(*
SPDX-FileCopyrightText: © 2026 Oleksandr Tiutyk <trofimich@gmail.com>
SPDX-License-Identifier: MIT
License: https://opensource.org/license/mit
*)

(*!
<summary>Provides shared comparer instances and selects them by generic value category.</summary>
<description>
Returned comparer interfaces borrow instances stored in this program; callers do not own or release them.
Selection does not inspect, validate or convert operand data. Callers must supply live descriptors whose
representations satisfy the selected concrete comparer. OBJECT selects natural ordering through IComparable;
it does not select byte or address ordering. Dictionary/set equality lookup is independent of this catalogue.
</description>
*)

PROGRAM StandardComparers
VAR_OUTPUT
	BoolComparer : BoolComparer;
	SIntComparer : SIntComparer;
	USIntComparer : USIntComparer;
	IntComparer : IntComparer;
	UIntComparer : UIntComparer;
	DIntComparer : DIntComparer;
	UDIntComparer : UDIntComparer;
	LIntComparer : LIntComparer;
	ULIntComparer : ULIntComparer;
	RealComparer : RealComparer;
	LRealComparer : LRealComparer;		
	StringComparer : StringComparer;
	WStringComparer : WStringComparer;
	TimeComparer : TimeComparer;
	LTimeComparer : LTimeComparer;
	DateComparer : DateComparer;
	LDateComparer : LDateComparer;
	DateAndTimeComparer : DateAndTimeComparer;
	LDateAndTimeComparer : LDateAndTimeComparer;
	TimeOfDayComparer : TimeOfDayComparer;	
	LTimeOfDayComparer : LTimeOfDayComparer;	
	ByteArrayComparer : ByteArrayComparer;
	ObjectComparer : ObjectComparer;
	//! <summary>Shared comparer that orders descriptor storage addresses without reading stored pointer values.</summary>
	StorageAddressComparer : StorageAddressComparer;	
END_VAR
VAR
	{attribute 'hide'} 
	_ClassName : STRING := __POUNAME();
END_VAR

{attribute 'monitoring' := 'call'}
PROPERTY ClassName : REFERENCE TO STRING
GET
ClassName REF= _ClassName;
END_GET
END_PROPERTY

(*!
<summary>Returns the shared comparer selected for a generic value category.</summary>
<description>
The result borrows a catalogue instance and does not transfer ownership. No operands are inspected or
converted; compatibility and operand lifetime remain the caller's responsibility. UNSPECIFIED and unknown
categories raise ArgumentOutOfRangeException. Concrete comparers define their supported representations and
null handling. OBJECT returns ObjectComparer, which uses IComparable for two non-null objects and rejects
missing natural-order support; USER_DEFINED retains byte ordering.
</description>
*)
//!<param name="typeClass">Generic representation category used to select the comparer.</param>
METHOD GetForTypeClass : TOF_Core.IComparer
VAR_INPUT
	typeClass : TOF_Core.GENERIC_TYPE_CLASS;
END_VAR
CASE typeClass OF
    TOF_Core.GENERIC_TYPE_CLASS.BOOLEAN:
		GetForTypeClass := BoolComparer;
    TOF_Core.GENERIC_TYPE_CLASS.INT_8:
		GetForTypeClass := SIntComparer;
    TOF_Core.GENERIC_TYPE_CLASS.INT_16:
		GetForTypeClass := IntComparer;
    TOF_Core.GENERIC_TYPE_CLASS.INT_32:
		GetForTypeClass := DIntComparer;
    TOF_Core.GENERIC_TYPE_CLASS.INT_64:
		GetForTypeClass := LIntComparer;
    TOF_Core.GENERIC_TYPE_CLASS.UINT_8:
		GetForTypeClass := USIntComparer;
    TOF_Core.GENERIC_TYPE_CLASS.UINT_16:
		GetForTypeClass := UIntComparer;
    TOF_Core.GENERIC_TYPE_CLASS.UINT_32:
		GetForTypeClass := UDIntComparer;
    TOF_Core.GENERIC_TYPE_CLASS.UINT_64:
		GetForTypeClass := ULIntComparer;
    TOF_Core.GENERIC_TYPE_CLASS.REAL_32:
		GetForTypeClass := RealComparer;
    TOF_Core.GENERIC_TYPE_CLASS.REAL_64:
		GetForTypeClass := LRealComparer;
    TOF_Core.GENERIC_TYPE_CLASS.STRING_8:
		GetForTypeClass := StringComparer;
    TOF_Core.GENERIC_TYPE_CLASS.STRING_16:
		GetForTypeClass := WStringComparer;
    TOF_Core.GENERIC_TYPE_CLASS.DATE_32:
		GetForTypeClass := DateComparer;
    TOF_Core.GENERIC_TYPE_CLASS.DATE_64:
		GetForTypeClass := LDateComparer;
    TOF_Core.GENERIC_TYPE_CLASS.TIME_32:
		GetForTypeClass := TimeComparer;
    TOF_Core.GENERIC_TYPE_CLASS.TIME_64:
		GetForTypeClass := LTimeComparer;
    TOF_Core.GENERIC_TYPE_CLASS.DATE_AND_TIME_32:
		GetForTypeClass := DateAndTimeComparer;
    TOF_Core.GENERIC_TYPE_CLASS.DATE_AND_TIME_64:
		GetForTypeClass := LDateAndTimeComparer;
    TOF_Core.GENERIC_TYPE_CLASS.TIME_OF_DAY_32:
		GetForTypeClass := TimeOfDayComparer;
    TOF_Core.GENERIC_TYPE_CLASS.TIME_OF_DAY_64:
		GetForTypeClass := LTimeOfDayComparer;
    TOF_Core.GENERIC_TYPE_CLASS.POINTER_TO:
		GetForTypeClass := StorageAddressComparer;
    TOF_Core.GENERIC_TYPE_CLASS.OBJECT:
		GetForTypeClass := ObjectComparer;
    TOF_Core.GENERIC_TYPE_CLASS.USER_DEFINED:
		GetForTypeClass := ByteArrayComparer;
	ELSE
		TOF_Core.Exceptions.ThrowArgumentOutOfRange(
			sourceNamespaceName := CurrentNamespace.Name,
			sourceClassName := ClassName,
			sourcePOUName := __POUNAME(),
			sourcePosition := __POSITION(),
			argumentName := 'typeClass',
			argumentValue := typeClass
		);
END_CASE
END_METHOD

(*!
<summary>Returns a borrowed read-only reference to this library's namespace name.</summary>
<description>
The storage belongs to CurrentNamespace and remains valid throughout the program instance lifetime.
</description>
*)
{attribute 'monitoring' := 'call'}
PROPERTY NamespaceName : REFERENCE TO STRING
GET
NamespaceName REF= CurrentNamespace.Name;
END_GET
END_PROPERTY

END_PROGRAM

(* stored: Version 1.1.0.1
   POU StandardComparers: Id {87b8ffe1-0355-4a7f-8d1d-1285b07f1992}, SpecialFunc None
   Property ClassName: Id {a555cabc-7156-4add-909f-9abd99c5db6a}
   Get Get: Id {57b1b255-8046-4561-b3ec-5fa164bac495}
   Method GetForTypeClass: Id {dc4a6532-4828-4b1a-a763-e1cc543032b4}
   Property NamespaceName: Id {8356e701-dddc-44e7-803f-9298ff48040a}
   Get Get: Id {e48cd34b-0adc-48ea-aa84-6f7122cba333} *)
